Staubli VAL3: updateInfo.pgx

public program updateInfo(num x_nItemIn, num& x_nItemOut, string& x_sTextOut, string x_sNo, string x_sComment)
  local string l_sTextOut
begin
  switch sLanguage
    case "chinese"
      l_sTextOut=sHmiCN[x_nItemIn]
    break
    case "english"
      l_sTextOut=sHmiEN[x_nItemIn]
    break
  endSwitch
  if x_sNo=="0" or x_nItemIn==100
    x_sTextOut=l_sTextOut
  else
    if x_nItemIn==99
      x_sTextOut=""
    else
      x_sTextOut=x_sNo+"."+l_sTextOut
    endIf
  endIf
  x_nItemOut=x_nItemIn
end
